// TIA Portal V19 export
TYPE "ST_TPM_AutoFeedback"
   STRUCT
      Ready : Bool;   // Ready to accept a new request (may fall while Busy).
      Busy : Bool;
      Done : Bool;
      Error : Bool;
      Aborted : Bool;
   END_STRUCT;
END_TYPE
